(* IEC 61131-3 sources: nautilus/website/lessons/b1-blink/variants/ok-nine-scans, 1 file *)

(* ---- program.st ---- *)
PROGRAM Blink
VAR n : INT; END_VAR
n := n + 1;
IF n >= 9 THEN
    Lamp := NOT Lamp;
    n := 0;
END_IF;
END_PROGRAM
